// TwinCAT 3 PLC project ueb_plc
// ProgramVersion: 3.1.4024.0
// libraries:
//   Tc2_EtherCAT, * (Beckhoff Automation GmbH)
//   Tc2_Standard, * (Beckhoff Automation GmbH)
//   Tc2_System, * (Beckhoff Automation GmbH)
//   Tc2_Utilities, * (Beckhoff Automation GmbH)
//   Tc3_EventLogger, * (Beckhoff Automation GmbH)
//   Tc3_Module, * (Beckhoff Automation GmbH)
// project tree:
//   GVLs/ GVL.TcGVL, GVL_InitEarly.TcGVL, GVL_InitLate.TcGVL
//   / PlcTask.TcTTO
//   POUs/ CD_Register.TcCD (not stored), FB_Base.TcPOU, FB_MyTimingSample.TcPOU, FB_MY_EVENT_MESSAGE.TcPOU, FB_Register.TcPOU, ITF_Base.TcIO, MAIN.TcPOU, PRG_AfterGlobalInit.TcPOU
// real-time tasks:
//   TASK PlcTask: cycle T#10ms, priority 20, ADS port 350

CONFIGURATION ueb_plc
    RESOURCE PLC ON TwinCAT3
        TASK PlcTask(INTERVAL := T#10ms, PRIORITY := 20);
        PROGRAM MAIN WITH PlcTask : MAIN;
    END_RESOURCE
END_CONFIGURATION

// ---- GVLs/GVL.TcGVL
{attribute 'qualified_only'}
{attribute 'global_init_slot' := '40001'}
VAR_GLOBAL
    Register : FB_REGISTER;
END_VAR

// ---- GVLs/GVL_InitEarly.TcGVL
{attribute 'qualified_only'}
{attribute 'global_init_slot' := '40001'}
VAR_GLOBAL
    nTimestamp : Tc2_EtherCAT.T_DCTIME64 :=
        Tc2_EtherCAT.F_GetActualDcTime64();
END_VAR

// ---- GVLs/GVL_InitLate.TcGVL
{attribute 'qualified_only'}
{attribute 'global_init_slot' := '59999'}
VAR_GLOBAL
    nTimestamp : Tc2_EtherCAT.T_DCTIME64 :=
        Tc2_EtherCAT.F_GetActualDcTime64();
END_VAR

// ---- POUs/ITF_Base.TcIO
INTERFACE ITF_Base

PROPERTY Error : UDINT
GET
END_GET
SET
END_SET
END_PROPERTY

END_INTERFACE

// ---- POUs/MAIN.TcPOU
PROGRAM MAIN
VAR
    fbMessage1 : FB_MY_EVENT_MESSAGE;
    fbMessage2 : FB_MY_EVENT_MESSAGE;

    nError1 : UDINT := 0;
    nError2 : UDINT := 0;

    sError1 : T_MaxString := 'Testfehler Wechselrichter';
    sError2 : T_MaxString := 'Testfehler Speicher';

    nNow : Tc2_EtherCAT.T_DCTIME64;
	
	fbTiming1 : FB_MyTimingSample;
	fbTiming2 : FB_MyTimingSample;
	
	fbBase1 : FB_Base;
    fbBase2 : FB_Base;
    fbBase3 : FB_Base;
	
	nErrorFromRegister : UDINT;
END_VAR

// Aktuelle DC-Zeit.
// Der Meldungsbaustein speichert sie beim Erkennen eines Fehlers.
nNow := Tc2_EtherCAT.F_GetCurDcTickTime64();

fbMessage1(
    sSourcename := 'Wechselrichter',
    eLevel     := Tc3_EventLogger.TcEventSeverity.Error,
    nEventCode := TC_EVENTS.EC_Uebungen.ExternalError.nEventId,
    nError     := nError1,
    sError     := sError1,
    nTimeStamp := nNow
);

fbMessage2(
    sSourcename := 'Speicher',
    eLevel     := Tc3_EventLogger.TcEventSeverity.Warning,
    nEventCode := TC_EVENTS.EC_Uebungen.ExternalError.nEventId,
    nError     := nError2,
    sError     := sError2,
    nTimeStamp := nNow
);

IF GVL.Register.arrRegister[1] <> 0 THEN
    nErrorFromRegister := GVL.Register.arrRegister[1].Error;
END_IF

END_PROGRAM

// ---- POUs/FB_MY_EVENT_MESSAGE.TcPOU
FUNCTION_BLOCK FB_MY_EVENT_MESSAGE
VAR_INPUT
    sSourcename : T_MaxString;
    eLevel     : Tc3_EventLogger.TcEventSeverity;
    nEventCode : UDINT;
    nError     : UDINT;
    sError     : T_MaxString;
    nTimeStamp : Tc2_EtherCAT.T_DCTIME64;
END_VAR

VAR
    fbTcSourceInfo : Tc3_EventLogger.FB_TcSourceInfo;
    fbTcMessage    : Tc3_EventLogger.FB_TcMessage;

    nStep          : UINT := 0;
    nLastError     : UDINT := 0;

    // Eingänge für die mehrzyklische Verarbeitung zwischenspeichern
    sSourceSaved   : T_MaxString;
    eLevelSaved    : Tc3_EventLogger.TcEventSeverity;
    nEventSaved    : UDINT;
    nErrorSaved    : UDINT;
    sErrorSaved    : T_MaxString;
    nTimeSaved     : Tc2_EtherCAT.T_DCTIME64;

    // Rückgabecode der EventLogger-Aufrufe
    hrResult       : HRESULT;
	
	nEventTime : ULINT;
END_VAR

CASE nStep OF

    0: // Änderung des Fehlercodes erkennen
        IF nError <> nLastError THEN
            // Auch den Wechsel auf 0 merken:
            // Derselbe Fehler kann danach erneut auftreten.
            nLastError := nError;

            IF nError > 0 THEN
                sSourceSaved := sSourcename;
                eLevelSaved  := eLevel;
                nEventSaved  := nEventCode;
                nErrorSaved  := nError;
                sErrorSaved  := sError;
                nTimeSaved   := nTimeStamp;

                nStep := 10;
            END_IF
        END_IF


    10: // Quelle setzen und Nachricht erstellen
        fbTcSourceInfo.Clear();
        fbTcSourceInfo.sName := sSourceSaved;

        hrResult := fbTcMessage.Create(
			eventClass   := TC_EVENTS.EC_Uebungen.ExternalError.uuidEventClass,
			nEventId     := nEventSaved,
			eSeverity    := eLevelSaved,
			ipSourceInfo := fbTcSourceInfo
		);
        IF hrResult = 0 THEN // S_OK
            nStep := 20;
        END_IF


    20: // Argumente setzen und Nachricht senden
        fbTcMessage.ipArguments.Clear();
        fbTcMessage.ipArguments.AddUDint(nErrorSaved);
        fbTcMessage.ipArguments.AddString(sErrorSaved);

        IF nTimeSaved = 0 THEN
            // Sonderfall: EventLogger verwendet die aktuelle Zeit.
            nEventTime := 0;
        ELSE
            nEventTime :=
                Tc2_EtherCAT.DCTIME64_TO_FILETIME64(nTimeSaved);
        END_IF

        hrResult := fbTcMessage.Send(
            nTimeStamp := nEventTime
        );

        IF hrResult = 0 THEN // S_OK
            nStep := 30;
        END_IF


    30: // Meldungsinstanz freigeben
        hrResult := fbTcMessage.Release();

        IF hrResult = 0 THEN // S_OK
            nStep := 0;
        END_IF

END_CASE

END_FUNCTION_BLOCK

// ---- POUs/FB_MyTimingSample.TcPOU
{attribute 'call_after_init'}
FUNCTION_BLOCK FB_MyTimingSample
VAR
    nTimestampFB_init   : Tc2_EtherCAT.T_DCTIME64;
    nTimestampFB_reinit : Tc2_EtherCAT.T_DCTIME64;
    nTimestampMyInit    : Tc2_EtherCAT.T_DCTIME64;
END_VAR

METHOD FB_init : BOOL
VAR_INPUT
    bInitRetains : BOOL;
    bInCopyCode  : BOOL;
END_VAR
nTimestampFB_init := Tc2_EtherCAT.F_GetActualDcTime64();
FB_init := TRUE;
END_METHOD

METHOD FB_reinit : BOOL
VAR_INPUT
END_VAR
nTimestampFB_reinit := Tc2_EtherCAT.F_GetActualDcTime64();
FB_reinit := TRUE;
END_METHOD

{attribute 'call_after_init'}
METHOD MyInit : BOOL
nTimestampMyInit := Tc2_EtherCAT.F_GetActualDcTime64();
MyInit := TRUE;
END_METHOD

END_FUNCTION_BLOCK

// ---- POUs/FB_Base.TcPOU
FUNCTION_BLOCK FB_Base IMPLEMENTS ITF_Base
VAR_INPUT
END_VAR
VAR_OUTPUT
END_VAR
VAR
	nErrorId     : UDINT := 0;
    nRegisterPos : UDINT := 0;
END_VAR

{warning 'Eigenschaftenimplementierung hinzufügen'}
PROPERTY Error : UDINT
GET
Error := nErrorId;
END_GET
SET
nErrorId := Error;
END_SET
END_PROPERTY

METHOD FB_init : BOOL
VAR_INPUT
	bInitRetains : BOOL; // if TRUE, the retain variables are initialized (warm start / cold start)
	bInCopyCode : BOOL;  // if TRUE, the instance afterwards gets moved into the copy code (online change)
END_VAR
nRegisterPos := GVL.Register.AddInterfacePointer(
    ipBase := THIS^
);

FB_init := TRUE;
END_METHOD

END_FUNCTION_BLOCK

// ---- POUs/FB_Register.TcPOU
FUNCTION_BLOCK FB_Register
VAR_INPUT
END_VAR
VAR_OUTPUT
END_VAR
VAR
	arrRegister     : ARRAY[1..100] OF ITF_Base;
    nNoOfInterfaces : UDINT := 0;
END_VAR

METHOD PUBLIC AddInterfacePointer : UDINT
VAR_INPUT
	ipBase : ITF_Base;
END_VAR
VAR
	n : UDINT;
END_VAR
// 0 bedeutet: Registrierung nicht erfolgreich.
AddInterfacePointer := 0;

// Eine leere Interface-Referenz nicht aufnehmen.
IF ipBase = 0 THEN
    RETURN;
END_IF

// Bereits registriert? Bestehenden Platz zurückgeben.
FOR n := 1 TO nNoOfInterfaces DO
    IF arrRegister[n] = ipBase THEN
        AddInterfacePointer := n;
        RETURN;
    END_IF
END_FOR

// Bei vollem Register nichts verändern.
IF nNoOfInterfaces >= 100 THEN
    RETURN;
END_IF

// Neue Referenz speichern.
nNoOfInterfaces := nNoOfInterfaces + 1;
arrRegister[nNoOfInterfaces] := ipBase;

// Zugewiesenen Tabellenplatz zurückgeben.
AddInterfacePointer := nNoOfInterfaces;
END_METHOD

END_FUNCTION_BLOCK

// ---- POUs/PRG_AfterGlobalInit.TcPOU
{attribute 'linkalways'}
{attribute 'call_after_global_init_slot' := '1'}
PROGRAM PRG_AfterGlobalInit
VAR
    nTimestampDeclaration : Tc2_EtherCAT.T_DCTIME64 :=
        Tc2_EtherCAT.F_GetActualDcTime64();

    nTimestampExecution : Tc2_EtherCAT.T_DCTIME64;
END_VAR

nTimestampExecution := Tc2_EtherCAT.F_GetActualDcTime64();

END_PROGRAM
